ABB RobotStudio station: Pallet_Project.rspag

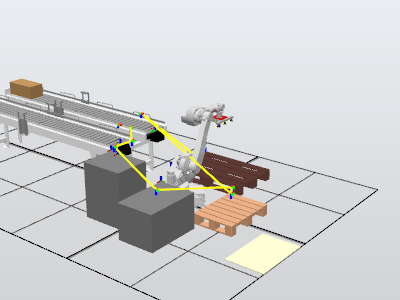
--- station ---
Station Pallet_Project (saved by RobotStudio 25.2.11220.0)
Controller Controler
  mechanical unit ROB_1: IRB1600_10_145__02, 6 joints, base frame (0, 0, 0) mm, rotated rx 0 ry 0 rz 135 deg
Layout (positions relative to the parent item):
  - IRB1600_10_145__02 [mechanism, from %ABB.RobotStudio.Models.IRB1600%\IRB1600_10_145_G_02.rslib] at (0, 0, 0) mm, rotated rx 0 ry 0 rz 135 deg; joint values [-2.2455, 0.5806, -0.4983, 0, 1.4885, 0.1107] (rad or m)
  - Half EPAL [part] at (-400, -600, 0) mm, rotated rx 0 ry 0 rz -90 deg, size 600 x 800 x 144 mm
  - ConveyorBox1 [part, from %ABB.RobotStudio.Models.Conveyors%\Conveyor Guide 400.rslib] at (150, 3660, 0) mm, rotated rx 0 ry 0 rz -90 deg
  - ConveyorBox2 [part, from %ABB.RobotStudio.Models.Conveyors%\Conveyor Guide 400.rslib] at (-550, 3660, 0) mm, rotated rx 0 ry 0 rz -90 deg
  - PalletizingVacuumTool [mechanism] at (1125, 125, 957.51) mm, rotated rx -180 ry 0 rz 180 deg
      TCP toolVacuum at (0, 0, 175) mm
      links: PalletizingVacuumTool
  - Box1 [part] at (338.5, 3410, 868) mm, size 249 x 499 x 200 mm
  - Box2 [part] at (-353.5, 3575, 868) mm, size 129 x 129 x 200 mm
  - EuroPallet [part, from Components\EuroPalletWood.rslib] at (1400, -600, 0) mm, rotated rx 0 ry 0 rz 90 deg
  - StackingTable [part], size 500 x 600 x 770 mm
  - LinerStand [part], size 800 x 540 x 500 mm
  - SC_Conveyor1 [smart component]
      signals: DO BoxArrived, DI EuroPalletReplaced, DO EuroPalletReplacedOut, DI EuroPalletFull
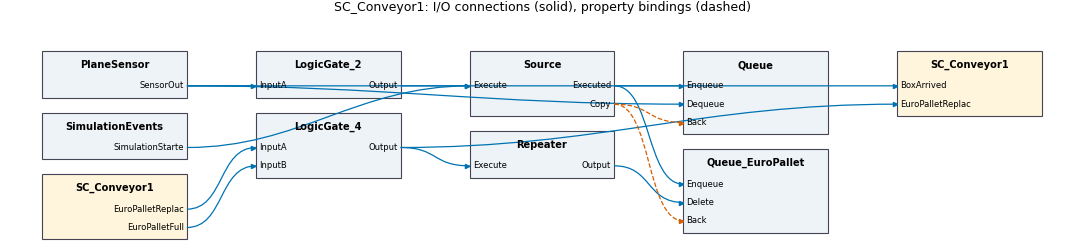
      connections:
        Source.Executed -> Queue.Enqueue
        PlaneSensor.SensorOut -> Queue.Dequeue
        PlaneSensor.SensorOut -> SC_Conveyor1.BoxArrived
        PlaneSensor.SensorOut -> LogicGate_2.InputA
        Source.Executed -> Queue_EuroPallet.Enqueue
        LogicGate_2.Output -> Source.Execute
        SimulationEvents.SimulationStarted -> Source.Execute
        SC_Conveyor1.EuroPalletReplaced -> LogicGate_4.InputA
        SC_Conveyor1.EuroPalletFull -> LogicGate_4.InputB
        LogicGate_4.Output -> Repeater.Execute
        LogicGate_4.Output -> SC_Conveyor1.EuroPalletReplacedOut
        Repeater.Output -> Queue_EuroPallet.Delete
        Source.Copy => Queue.Back
        Source.Copy => Queue_EuroPallet.Back
    - Source [smart component, from Components\Source.rslib]
        properties: Source=Box1; Copy=(none); Parent=(none); Position=[0.3385 3.39 0.868]; Orientation=[0 0 0]; Transient=true; PhysicsBehavior=-1
    - Queue [smart component, from Components\Queue.rslib]
        properties: Back=(none); Front=(none); Queue={81e52df3-1f77-4299-ba2a-6414327be985};{435d0d6d-d79b-44d3-acea-fe52ef949857};{8436b295-f8bf-4107-9481-0b8da08c6045};{6da8449d-009c-4835-8de1-a31c03bf24d8};{c517003d-8767-4c4a-bff9-7cbe8e804e1a};{f09c25fa-2584-409c-84e2-e14a50677c13};{130e9f86-ac44-4070-b92e-1e55d896aa7b};{906d2277-e14e-41d7-b5ad-7fe71654f1ef};{c971c019-2e6c-4537-9b43-f56770b68a66};{5740a0fa-eee5-4cb0-a52c-79e90074768b};{0e505042-845a-40e7-8904-6deb6f228de7};{2ef81a46-8090-4cc3-a468-447f4544bad1};{dd80a3b0-d0cd-4f2f-9600-d92ba7686845};{3b519026-604d-4377-8cfe-ae9118f60529}; NumberOfObjects=1
    - LinearMover [smart component, from Components\LinearMover.rslib]
        properties: Object=Queue; Direction=[0 -0.001 0]; Speed=0.25; Reference=Global; ReferenceObject=(none)
    - PlaneSensor [smart component, from Components\PlaneSensor.rslib]
        properties: Origin=[0.1885 0.675 0.788]; Axis1=[0.3 0 0]; Axis2=[0 0 0.01]; Tag=(none); SenseMultiple=false; SensedPart=(none)
      - _sensorPart_ [part], size 300 x 0 x 10 mm
    - LogicGate_2 [smart component, from Components\LogicGate.rslib]
        properties: Operator=NOT; Delay=0
    - SimulationEvents [smart component, from Components\SimulationEvents.rslib]
    - Queue_EuroPallet [smart component, from Components\Queue.rslib]
        properties: Back=(none); Front=(none); Queue={2ef81a46-8090-4cc3-a468-447f4544bad1};{dd80a3b0-d0cd-4f2f-9600-d92ba7686845};{3b519026-604d-4377-8cfe-ae9118f60529}; NumberOfObjects=3
    - LogicGate_4 [smart component, from Components\LogicGate.rslib]
        properties: Operator=AND; Delay=0
    - Repeater [smart component, from Components\Repeater.rslib]
        properties: Count=12
  - SC_Gripper [smart component]
      signals: DI Grip
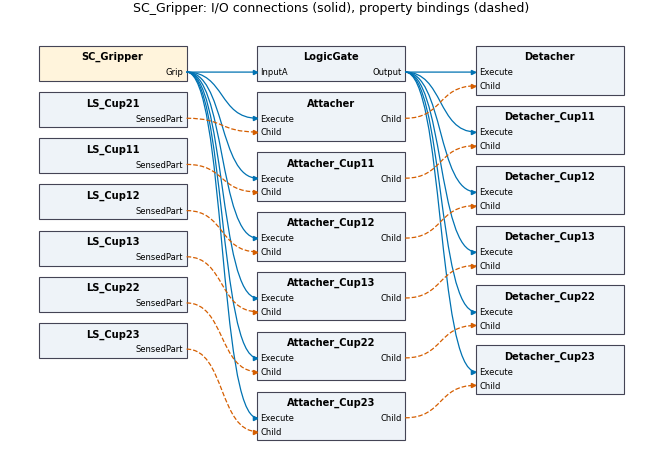
      connections:
        SC_Gripper.Grip -> Attacher.Execute
        SC_Gripper.Grip -> LogicGate.InputA
        LogicGate.Output -> Detacher.Execute
        SC_Gripper.Grip -> Attacher_Cup11.Execute
        LogicGate.Output -> Detacher_Cup11.Execute
        SC_Gripper.Grip -> Attacher_Cup12.Execute
        LogicGate.Output -> Detacher_Cup12.Execute
        SC_Gripper.Grip -> Attacher_Cup13.Execute
        LogicGate.Output -> Detacher_Cup13.Execute
        SC_Gripper.Grip -> Attacher_Cup22.Execute
        LogicGate.Output -> Detacher_Cup22.Execute
        SC_Gripper.Grip -> Attacher_Cup23.Execute
        LogicGate.Output -> Detacher_Cup23.Execute
        LS_Cup21.SensedPart => Attacher.Child
        Attacher.Child => Detacher.Child
        LS_Cup11.SensedPart => Attacher_Cup11.Child
        Attacher_Cup11.Child => Detacher_Cup11.Child
        LS_Cup12.SensedPart => Attacher_Cup12.Child
        Attacher_Cup12.Child => Detacher_Cup12.Child
        LS_Cup13.SensedPart => Attacher_Cup13.Child
        Attacher_Cup13.Child => Detacher_Cup13.Child
        LS_Cup22.SensedPart => Attacher_Cup22.Child
        Attacher_Cup22.Child => Detacher_Cup22.Child
        LS_Cup23.SensedPart => Attacher_Cup23.Child
        Attacher_Cup23.Child => Detacher_Cup23.Child
    - LS_Cup21 [smart component, from Components\LineSensor.rslib] at (375, 125, -163.99) mm, rotated rx 0 ry 0 rz -135 deg
        properties: Start=[-0.597509982704304 0.689429996191639 0.956499992313755]; End=[-0.597509981617333 0.689429995104668 0.924499992313755]; Length=0.032; Radius=0.00331491712707182; Tag=(none); SenseMultiple=false; SensedPart=(none); SensedPoint=[0 0 0]
      - _sensorPart_ [part], size 6.4 x 6.4 x 32 mm
    - Attacher [smart component, from Components\Attacher.rslib]
        properties: Parent=PalletizingVacuumTool; Flange=0; Child=(none); Mount=false; Offset=[0 0 0]; Orientation=[0 0 0]
    - Detacher [smart component, from Components\Detacher.rslib]
        properties: Child=(none); KeepPosition=true
    - LogicGate [smart component, from Components\LogicGate.rslib]
        properties: Operator=NOT; Delay=0
    - LS_Cup11 [smart component, from Components\LineSensor.rslib] at (375, 125, -163.99) mm, rotated rx 0 ry 0 rz -135 deg
        properties: Start=[-0.68943 0.59751 0.9565]; End=[-0.68943 0.59751 0.9245]; Length=0.032; Radius=0.00331; Tag=(none); SenseMultiple=false; SensedPart=(none); SensedPoint=[0 0 0]
      - _sensorPart_ [part], size 6.6 x 6.6 x 32 mm
    - LS_Cup12 [smart component, from Components\LineSensor.rslib] at (375, 125, -163.99) mm, rotated rx 0 ry 0 rz -135 deg
        properties: Start=[-0.57629 0.48437 0.9565]; End=[-0.57629 0.48437 0.9245]; Length=0.032; Radius=0.00331; Tag=(none); SenseMultiple=false; SensedPart=(none); SensedPoint=[0 0 0]
      - _sensorPart_ [part], size 6.6 x 6.6 x 32 mm
    - LS_Cup13 [smart component, from Components\LineSensor.rslib] at (375, 125, -163.99) mm, rotated rx 0 ry 0 rz -135 deg
        properties: Start=[-0.46315 0.37123 0.9565]; End=[-0.46315 0.37123 0.9245]; Length=0.032; Radius=0.00331; Tag=(none); SenseMultiple=false; SensedPart=(none); SensedPoint=[0 0 0]
      - _sensorPart_ [part], size 6.6 x 6.6 x 32 mm
    - LS_Cup22 [smart component, from Components\LineSensor.rslib] at (375, 125, -163.99) mm, rotated rx 0 ry 0 rz -135 deg
        properties: Start=[-0.48437 0.57629 0.9565]; End=[-0.48437 0.57629 0.9245]; Length=0.032; Radius=0.00331; Tag=(none); SenseMultiple=false; SensedPart=(none); SensedPoint=[0 0 0]
      - _sensorPart_ [part], size 6.6 x 6.6 x 32 mm
    - LS_Cup23 [smart component, from Components\LineSensor.rslib] at (375, 125, -163.99) mm, rotated rx 0 ry 0 rz -135 deg
        properties: Start=[-0.37123 0.46315 0.9565]; End=[-0.37123 0.46315 0.9245]; Length=0.032; Radius=0.00331; Tag=(none); SenseMultiple=false; SensedPart=(none); SensedPoint=[0 0 0]
      - _sensorPart_ [part], size 6.6 x 6.6 x 32 mm
    - Attacher_Cup11 [smart component, from Components\Attacher.rslib]
        properties: Parent=PalletizingVacuumTool; Flange=0; Child=(none); Mount=false; Offset=[0 0 0]; Orientation=[0 0 0]
    - Detacher_Cup11 [smart component, from Components\Detacher.rslib]
        properties: Child=(none); KeepPosition=true
    - Attacher_Cup12 [smart component, from Components\Attacher.rslib]
        properties: Parent=PalletizingVacuumTool; Flange=0; Child=(none); Mount=false; Offset=[0 0 0]; Orientation=[0 0 0]
    - Detacher_Cup12 [smart component, from Components\Detacher.rslib]
        properties: Child=(none); KeepPosition=true
    - Attacher_Cup13 [smart component, from Components\Attacher.rslib]
        properties: Parent=PalletizingVacuumTool; Flange=0; Child=(none); Mount=false; Offset=[0 0 0]; Orientation=[0 0 0]
    - Detacher_Cup13 [smart component, from Components\Detacher.rslib]
        properties: Child=(none); KeepPosition=true
    - Attacher_Cup22 [smart component, from Components\Attacher.rslib]
        properties: Parent=PalletizingVacuumTool; Flange=0; Child=(none); Mount=false; Offset=[0 0 0]; Orientation=[0 0 0]
    - Detacher_Cup22 [smart component, from Components\Detacher.rslib]
        properties: Child=(none); KeepPosition=true
    - Attacher_Cup23 [smart component, from Components\Attacher.rslib]
        properties: Parent=PalletizingVacuumTool; Flange=0; Child=(none); Mount=false; Offset=[0 0 0]; Orientation=[0 0 0]
    - Detacher_Cup23 [smart component, from Components\Detacher.rslib]
        properties: Child=(none); KeepPosition=true
  - SC_Conveyor2 [smart component]
      signals: DO BoxArrived, DI HalfPalletReplaced, DI HalfPalletFull, DO HalfPalletReplacedOut
      connections:
        Source.Executed -> Queue.Enqueue
        PlaneSensor.SensorOut -> Queue.Dequeue
        PlaneSensor.SensorOut -> SC_Conveyor2.BoxArrived
        PlaneSensor.SensorOut -> LogicGate.InputA
        SimulationEvents.SimulationStarted -> Source.Execute
        LogicGate.Output -> Source.Execute
        Repeater.Output -> Queue_HalfPallet.Delete
        SC_Conveyor2.HalfPalletReplaced -> LogicGate_5.InputA
        SC_Conveyor2.HalfPalletFull -> LogicGate_5.InputB
        LogicGate_5.Output -> Repeater.Execute
        LogicGate_5.Output -> SC_Conveyor2.HalfPalletReplacedOut
        Source.Executed -> Queue_HalfPallet.Enqueue
        Source.Copy => Queue.Back
        Source.Copy => Queue_HalfPallet.Back
    - Source [smart component, from Components\Source.rslib]
        properties: Source=Box2; Copy=(none); Parent=(none); Position=[-0.3535 3.575 0.868]; Orientation=[0 0 0]; Transient=true; PhysicsBehavior=-1
    - Queue [smart component, from Components\Queue.rslib]
        properties: Back=(none); Front=(none); Queue={9800cfb8-accd-4327-91e1-8f1786e05042};{c190d427-2878-4db8-b2be-214c692a7843};{b2a63077-10cd-4047-b774-a402e54bd5ce};{0cb034eb-9137-4204-8c4d-aa4d35edbbb2};{a2136454-01e3-48eb-803c-0c949220dd1f};{d1d29149-a959-4839-a5f8-05156c3e548d};{48c194bf-a44f-484f-bd23-34306ecfb550};{495763de-9b16-4c8d-83d3-4557bdb480a3};{abf2df07-53cd-488b-8dcb-fd67f1eb4dba}; NumberOfObjects=0
    - LinearMover [smart component, from Components\LinearMover.rslib]
        properties: Object=Queue; Direction=[0 -0.001 0]; Speed=0.25; Reference=Global; ReferenceObject=(none)
    - PlaneSensor [smart component, from Components\PlaneSensor.rslib]
        properties: Origin=[-0.5035 0.675 0.788]; Axis1=[0.3 0 0]; Axis2=[0 0 0.01]; Tag=(none); SenseMultiple=false; SensedPart=(none)
      - _sensorPart_ [part], size 300 x 0 x 10 mm
    - LogicGate [smart component, from Components\LogicGate.rslib]
        properties: Operator=NOT; Delay=0
    - SimulationEvents [smart component, from Components\SimulationEvents.rslib]
    - Queue_HalfPallet [smart component, from Components\Queue.rslib]
        properties: Back=(none); Front=(none); Queue={d5a67242-ef94-4595-a834-178362eb1d62};{353021ae-f387-47f5-aad2-fe3f1426ad48};{d78ca7a8-fd6f-498f-a8d6-0ea3578c76b0};{3356f02f-29aa-44c2-9ebf-5d29c5a600e5};{8f4d4553-4c1d-4056-aeb8-bca03c426780};{1a6d2d73-c05b-4390-90bb-4172aa34495b};{5c83e94b-c9dd-45e1-939f-1611cce13607};{08b3fadb-cba7-4510-a02f-3e66ae7e4329};{3ef4086a-d1f9-4a83-9755-3951cf9eaa00};{7bbd94bd-538e-428e-af81-32894a937116};{23a64fb5-90dc-4163-9a5d-a709f29cb737};{65ed0540-bcad-4628-84d7-59a3b9c76640};{b98fc11a-8ded-4a1c-bcf2-f2c76b1d1bd5};{5eac1296-3e35-4c81-a158-90d5fa5352fe};{05c4dc44-4e6c-4dc2-9677-a1940e3b3e4c};{d3d90d6c-55f3-41f9-ab59-03e6f986434c};{de9bd2e6-7614-4944-a633-7d4466c06302};{d5320c6f-757c-466b-aded-364807c4b01e};{23621476-4bd4-41d2-9f29-d7724955c74c};{817a93c2-45d8-40d3-ae92-600157ce3ee9};{243d6776-53f3-40e8-a26d-04ab6a776894};{7c17ee41-3d5e-4ce3-b2c1-8319b1484f6c};{7a467470-9a85-48d0-bfc9-40585f186b4a};{7fbfd87a-23fa-474d-b93a-b31788b7d83a};{49c53e7e-6fec-4cf6-ade2-eccfaa663d3f};{fd420bc1-af1d-47a6-a241-17656bc699f2};{1442cd0c-dbcc-4cc3-9371-290095dab2c2};{d4afd0ce-8611-4c71-934e-ce83a9ed8ab0};{4a599a5b-b82c-4c22-8dc8-b659788bcb6c};{af434e4d-6f74-4bd4-92e4-29d48b0c2391};{1d1a6925-ca0b-4280-b7e3-c3d429ecdeb1};{5f6f7c8a-25f7-4961-bc3d-06f26c3590e9};{0a446cc8-67bf-4709-be5a-1f56f3673959};{1af88ff7-cf78-4e6d-9326-b5fe289dfe55};{5a76c50a-250b-45d0-bcc3-a15c7678bea9};{ce2ad899-ab0c-4e8d-b6d7-b5ce0875e251};{41250e61-ba51-4579-939a-c1cb9538416c};{f048b52f-5fa1-4572-b32f-60b2a46e1837};{1087fd67-f502-4529-85a7-08891c247a62};{a8fcad14-50a7-40f1-a4f5-1777183cc2f1};{093bf0cb-478b-4d41-bc85-a01e6c4947d5};{ba12b4d4-5356-412c-9a5b-07d0d090cd25};{ef8538f7-904e-4b24-81ca-ce6b8f30748f};{1e7db033-e1a6-46cf-8960-0a3b92aa4569};{6ae3754e-0c7d-46a2-8cb0-0df03192a8af};{a9820d8c-191d-4cb3-b284-618a32150a08};{67edf359-12bc-49fc-a518-7b7d3cdaf041};{ad25e574-dc3f-4262-b019-213ebc35634b};{9ab4d7b7-70db-4a3c-b7ba-4ffa764225eb};{e3a4e5db-fe34-4e2c-bab2-f43d24e1bbe5};{2af16a20-02e3-4091-b49e-02ac578eafb8};{1fd54043-75f1-4856-9dc4-5fcdc28b2d30};{b3ff0692-c2c4-465f-bc5c-501c830a156d};{c5881555-d748-47b7-88bf-bb4395c5d677};{22d02747-187f-42da-b66b-aeac508d4faf};{4d19efbb-6ba8-4530-9818-c3b36a5b5e6d};{c26dfd74-1de5-480f-8d87-a956ac996da4};{800d2495-1f8a-4fba-a20e-307d73ad8d62};{4b542189-3f8e-408f-9294-fa7737ba2a1e};{b91039b3-272a-456d-b4ad-0c586638a480};{a02115cb-f377-4e0b-9fca-d98f58ac551d};{4b29cf1c-701e-48c2-bed8-74150284ae2a};{1a79b9b6-686e-4284-baae-745627c15955};{ca69f178-3ff4-4429-a57f-e75714190848};{2eeff9d0-5db0-4a2e-8983-6baf0d7612ee};{eb15173f-71b9-4843-b116-0fef5b8487ca};{f03858ea-60b5-4441-9128-abbe714a5bd1};{88a7fade-b898-403a-9912-eb07dfa3f617};{0c60aaed-4d54-4bbc-a941-b06aadfbebd1};{9800cfb8-accd-4327-91e1-8f1786e05042};{c190d427-2878-4db8-b2be-214c692a7843};{b2a63077-10cd-4047-b774-a402e54bd5ce};{0cb034eb-9137-4204-8c4d-aa4d35edbbb2};{a2136454-01e3-48eb-803c-0c949220dd1f};{d1d29149-a959-4839-a5f8-05156c3e548d};{48c194bf-a44f-484f-bd23-34306ecfb550};{495763de-9b16-4c8d-83d3-4557bdb480a3};{abf2df07-53cd-488b-8dcb-fd67f1eb4dba}; NumberOfObjects=32
    - Repeater [smart component, from Components\Repeater.rslib]
        properties: Count=72
    - LogicGate_5 [smart component, from Components\LogicGate.rslib]
        properties: Operator=AND; Delay=0
  - Liner_01 [part] at (-900, -2000, 0) mm, size 800 x 540 x 10 mm
  - SC_Liners [smart component]
      signals: DI LinersRefilled, DI LinerStackEmpty, DI PalletReplaced, DO LinersRefilledOut
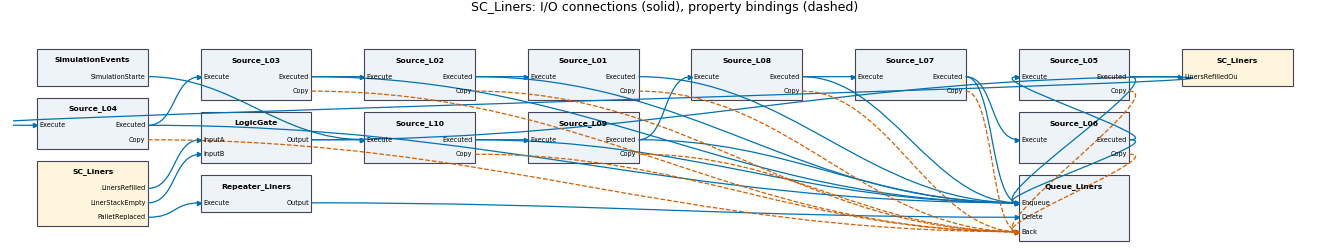
      connections:
        SimulationEvents.SimulationStarted -> Source_L10.Execute
        Source_L10.Executed -> Queue_Liners.Enqueue
        Source_L10.Executed -> Source_L09.Execute
        Source_L09.Executed -> Queue_Liners.Enqueue
        Source_L09.Executed -> Source_L08.Execute
        Source_L08.Executed -> Queue_Liners.Enqueue
        Source_L08.Executed -> Source_L07.Execute
        Source_L07.Executed -> Queue_Liners.Enqueue
        Source_L07.Executed -> Source_L06.Execute
        Source_L06.Executed -> Queue_Liners.Enqueue
        Source_L06.Executed -> Source_L05.Execute
        Source_L05.Executed -> Queue_Liners.Enqueue
        Source_L05.Executed -> Source_L04.Execute
        Source_L04.Executed -> Queue_Liners.Enqueue
        Source_L04.Executed -> Source_L03.Execute
        Source_L03.Executed -> Queue_Liners.Enqueue
        Source_L03.Executed -> Source_L02.Execute
        Source_L02.Executed -> Queue_Liners.Enqueue
        Source_L02.Executed -> Source_L01.Execute
        Source_L01.Executed -> Queue_Liners.Enqueue
        SC_Liners.LinersRefilled -> LogicGate.InputA
        SC_Liners.LinerStackEmpty -> LogicGate.InputB
        LogicGate.Output -> SC_Liners.LinersRefilledOut
        LogicGate.Output -> Source_L10.Execute
        SC_Liners.PalletReplaced -> Repeater_Liners.Execute
        Repeater_Liners.Output -> Queue_Liners.Delete
        Source_L10.Copy => Queue_Liners.Back
        Source_L09.Copy => Queue_Liners.Back
        Source_L08.Copy => Queue_Liners.Back
        Source_L07.Copy => Queue_Liners.Back
        Source_L06.Copy => Queue_Liners.Back
        Source_L05.Copy => Queue_Liners.Back
        Source_L04.Copy => Queue_Liners.Back
        Source_L03.Copy => Queue_Liners.Back
        Source_L02.Copy => Queue_Liners.Back
        Source_L01.Copy => Queue_Liners.Back
    - Source_L10 [smart component, from Components\Source.rslib]
        properties: Source=Liner_01; Copy=(none); Parent=(none); Position=[-1.3 -0.7 0.59]; Orientation=[0 0 0]; Transient=true; PhysicsBehavior=-1
    - Source_L09 [smart component, from Components\Source.rslib]
        properties: Source=Liner_01; Copy=(none); Parent=(none); Position=[-1.3 -0.7 0.58]; Orientation=[0 0 0]; Transient=true; PhysicsBehavior=-1
    - Queue_Liners [smart component, from Components\Queue.rslib]
        properties: Back=(none); Front=(none); Queue={20d974b6-189e-48d5-91a3-27801e75a2e3};{290c2d17-6faa-4c17-875c-80c899971b7e};{09f81150-e011-45c7-9a87-29c6d5ac92f7};{b296464f-7b57-4359-8933-3b585c425c6c};{a4bcdc79-e721-4592-ba3d-6f160afd2660};{d0cb2024-c7d0-4f62-9559-4447ca439c63};{f1537fa3-356e-4cfb-b79c-b3a3ef2d5a1a};{ade4e0be-57dc-4cbd-9040-6b29c36965ae};{068dc0fe-76cb-4174-b384-f9a97e7185e6};{74ebf040-bda5-45b9-9c71-05d8b50facaf};{455b281d-0163-4b9a-96ec-b3dbceeb94ec};{5721ff76-6329-4602-9dd2-421615ef1c3b}; NumberOfObjects=10
    - SimulationEvents [smart component, from Components\SimulationEvents.rslib]
    - Source_L08 [smart component, from Components\Source.rslib]
        properties: Source=Liner_01; Copy=(none); Parent=(none); Position=[-1.3 -0.7 0.57]; Orientation=[0 0 0]; Transient=true; PhysicsBehavior=-1
    - Source_L07 [smart component, from Components\Source.rslib]
        properties: Source=Liner_01; Copy=(none); Parent=(none); Position=[-1.3 -0.7 0.56]; Orientation=[0 0 0]; Transient=true; PhysicsBehavior=-1
    - Source_L06 [smart component, from Components\Source.rslib]
        properties: Source=Liner_01; Copy=(none); Parent=(none); Position=[-1.3 -0.7 0.55]; Orientation=[0 0 0]; Transient=true; PhysicsBehavior=-1
    - Source_L05 [smart component, from Components\Source.rslib]
        properties: Source=Liner_01; Copy=(none); Parent=(none); Position=[-1.3 -0.7 0.54]; Orientation=[0 0 0]; Transient=true; PhysicsBehavior=-1
    - Source_L04 [smart component, from Components\Source.rslib]
        properties: Source=Liner_01; Copy=(none); Parent=(none); Position=[-1.3 -0.7 0.53]; Orientation=[0 0 0]; Transient=true; PhysicsBehavior=-1
    - Source_L03 [smart component, from Components\Source.rslib]
        properties: Source=Liner_01; Copy=(none); Parent=(none); Position=[-1.3 -0.7 0.52]; Orientation=[0 0 0]; Transient=true; PhysicsBehavior=-1
    - Source_L02 [smart component, from Components\Source.rslib]
        properties: Source=Liner_01; Copy=(none); Parent=(none); Position=[-1.3 -0.7 0.51]; Orientation=[0 0 0]; Transient=true; PhysicsBehavior=-1
    - Source_L01 [smart component, from Components\Source.rslib]
        properties: Source=Liner_01; Copy=(none); Parent=(none); Position=[-1.3 -0.7 0.5]; Orientation=[0 0 0]; Transient=true; PhysicsBehavior=-1
    - LogicGate [smart component, from Components\LogicGate.rslib]
        properties: Operator=AND; Delay=0
    - Repeater_Liners [smart component, from Components\Repeater.rslib]
        properties: Count=2
Attachment: PalletizingVacuumTool is attached to IRB1600_10_145__02 / Link6
Attachment: LS_Cup21 is attached to PalletizingVacuumTool / PalletizingVacuumTool
Attachment: LS_Cup12 is attached to PalletizingVacuumTool / PalletizingVacuumTool
Attachment: LS_Cup13 is attached to PalletizingVacuumTool / PalletizingVacuumTool
Attachment: LS_Cup22 is attached to PalletizingVacuumTool / PalletizingVacuumTool
Attachment: LS_Cup23 is attached to PalletizingVacuumTool / PalletizingVacuumTool
Attachment: LS_Cup11 is attached to PalletizingVacuumTool / PalletizingVacuumTool
Collision set Conjunto de colisión_1: IRB1600_10_145__02, PalletizingVacuumTool against ConveyorBox1, ConveyorBox2, EuroPallet, Half EPAL, LinerStand, StackingTable, near miss 0.05 m
Station logic (signal -> signal, property => property):
  SC_Conveyor1.BoxArrived -> Controler.DI_Box1Arrived
  Controler.DO_Cup21 -> SC_Gripper.Grip
  SC_Conveyor2.BoxArrived -> Controler.DI_Box2Arrived
  SC_Conveyor1.EuroPalletReplacedOut -> Controler.DI_EuroPalletReplaced
  Controler.DO_EuroPalletFull -> SC_Conveyor1.EuroPalletFull
  Controler.DO_HalfPalletFull -> SC_Conveyor2.HalfPalletFull
  SC_Conveyor2.HalfPalletReplacedOut -> Controler.DI_HalfPalletReplaced
  Controler.DO_LinerStackEmpty -> SC_Liners.LinerStackEmpty
  SC_Liners.LinersRefilledOut -> Controler.DI_LinersRefilled
  SC_Conveyor2.HalfPalletReplacedOut -> SC_Liners.PalletReplaced
Targets, tools, work objects and paths stored in the station and not in the controller backup, written as RAPID:
! task T_ROB1
MODULE PalletProgram
  PROC Path_10()
    MoveL PickConveyor2,v1000,z100,toolVacuum\WObj:=wobjConveyor2;
    MoveL PlaceTable,v1000,z100,toolVacuum\WObj:=wobjTable;
    MoveL PickTableStack,v1000,z100,toolVacuum\WObj:=wobjTable;
    MoveL PickLiner,v1000,z100,toolVacuum\WObj:=wobjLinerStack;
    MoveL PlaceHalfPallet,v1000,z100,toolVacuum\WObj:=wobjHalfPallet;
    MoveL PlaceLiner,v1000,z100,toolVacuum\WObj:=wobjHalfPallet;
    MoveL PickConveyor1,v1000,z100,toolVacuum\WObj:=wobjConveyor1;
    MoveL PlaceEuroRow2,v1000,z100,toolVacuum\WObj:=wobjEuroPallet;
    MoveL PlaceEuroRow4,v1000,z100,toolVacuum\WObj:=wobjEuroPallet;
  ENDPROC
ENDMODULE


--- Controller Data/Controler/RAPID/TASK1/PROGMOD/CalibData.mod ---
MODULE CalibData
    !-----------------------------------------------------------------------
	! Tools and work object
	!-----------------------------------------------------------------------
    TASK PERS wobjdata wobjEuroPallet:=[FALSE,TRUE,"",[[600,600,144],[0.707106781,0,0,-0.707106781]],[[0,0,0],[1,0,0,0]]];
    TASK PERS wobjdata wobjHalfPallet:=[FALSE,TRUE,"",[[400,-600,144],[0,0,0,1]],[[0,0,0],[1,0,0,0]]];
    TASK PERS wobjdata wobjConveyor1:=[FALSE,TRUE,"",[[338.5,670,768],[0.707106781,0,0,0.707106781]],[[0,0,0],[1,0,0,0]]];
    TASK PERS wobjdata wobjConveyor2:=[FALSE,TRUE,"",[[-353.5,670,768],[0.707106781,0,0,0.707106781]],[[0,0,0],[1,0,0,0]]];
    TASK PERS wobjdata wobjTable:=[FALSE,TRUE,"",[[-600,600,770],[0,0,0,1]],[[55,170,0],[1,0,0,0]]];
    TASK PERS wobjdata wobjLinerStack:=[FALSE,TRUE,"",[[-500,-160,500],[0,0,0,1]],[[0,0,0],[1,0,0,0]]];
    TASK PERS tooldata toolVacuum:=[TRUE,[[0,0,175],[1,0,0,0]],[1,[0,0,1],[1,0,0,0],0,0,0]];
    ! toolVacuum: mass and CoG are provisional (1 kg), to be estimated

    !-----------------------------------------------------------------------
	! Load data
	!-----------------------------------------------------------------------
    ! Payloads: CoG relative to the TCP of toolVacuum; inertia set to 0 (point mass) until confirmed
    TASK PERS loaddata loadBox1:=[2,[0,0,100],[1,0,0,0],0,0,0];
    ! Box 2 is picked with one corner cup (x=-160, y=-100); on the table fill rows ascending Y, each row descending X
    TASK PERS loaddata loadBox2:=[0.4,[-160,-100,100],[1,0,0,0],0,0,0];
    ! 3x2 stack of box 2 (390 x 260 x 200 mm, 6 x 0.4 kg)
    TASK PERS loaddata loadBox2Stack:=[2.4,[0,0,100],[1,0,0,0],0,0,0];
    ! Liner: corrugated cardboard, 0.8 x 0.54 x 0.01 m3 x 120 kg/m3 = 0.52 kg
    TASK PERS loaddata loadLiner:=[0.52,[0,0,5],[1,0,0,0],0,0,0];
ENDMODULE

--- Controller Data/Controler/RAPID/TASK1/PROGMOD/PalletProgram.mod ---
MODULE PalletProgram

    !***********************************************************************
    ! Industrial Robotics and Offline Programming G1F - University of Skovde
    ! Offline programming project: Pallet Project - Group 2 (JMPM)
    ! Authors: Peru Mendivil and Joaquin Moreno
    ! Robot :   ABB IRB 1600-10/1.45, IRC5 RobotWare 6.13.02 (RobotStudio 2025)
    ! Tool  :   toolVacuum, vacuum gripper with 6 cups (one valve per cup)
    ! Date:    2026-10-30
    !
    ! The robot palletizes two products coming on two conveyors.
    ! Box 1 goes from conveyor 1 to the Euro pallet: 4-2 pattern,
    ! 2 layers (12 boxes). Box 2 goes from conveyor 2 to the stacking
    ! table, where a 3x2 block is formed. The block is then moved to the
    ! half pallet: 2x2 blocks per layer, 3 layers (72 boxes), with a liner
    ! after layers 1 and 2. When both conveyors have a box, the robot
    ! alternates box 1 and box 2. A full pallet is replaced by the operator
    ! from outside the fence, and the robot keeps working with the other
    ! product. With the half pallet full, one block can still be finished
    ! on the table, and it waits there. If the liner stack is empty, the
    ! robot keeps working until a liner is needed; then box 2 waits until
    ! the operator refills the stack.
    !
    ! Structure: Main is a state machine (grafcet). It initialises the
    ! signals and then decides each cycle which box to handle, from the
    ! conveyor sensors, the full-pallet flags and the last box handled.
    ! Each product has its own routine with a finite-state machine for
    ! the place positions. Every place position is calculated with Offs
    ! from one base target per station. ApproachPoint does every
    ! pick/place: approach, vacuum on/off and GripLoad. Work objects,
    ! tool and loads are in the module CalibData.
    ! The operator buttons (pallet replaced, liners refilled) are read
    ! with interrupts (TRAP), so a short press is never lost.
    !
    ! Naming: VAR, PERS and parameters in camelCase (can change);
    ! CONST, PROC, FUNC and MODULE in PascalCase (fixed).
    !***********************************************************************

    !-----------------------------------------------------------------------
    ! Base targets
    !-----------------------------------------------------------------------
    CONST jointtarget Home:=[[0,0,0,0,90,0],[9E+09,9E+09,9E+09,9E+09,9E+09,9E+09]];

    ! Box 1
    CONST robtarget PickConveyor1:=[[249.5,0,200],[0,0,1,0],[0,0,0,0],[9E+09,9E+09,9E+09,9E+09,9E+09,9E+09]];
    CONST robtarget PlaceEuroRow4:=[[225,525,200],[0,-0.707106781,0.707106781,0],[-2,0,0,0],[9E+09,9E+09,9E+09,9E+09,9E+09,9E+09]];
    CONST robtarget PlaceEuroRow2:=[[350,150,200],[0,1,0,0],[-2,0,-1,0],[9E+09,9E+09,9E+09,9E+09,9E+09,9E+09]];

    ! Box 2
    CONST robtarget PickConveyor2:=[[-35.5,-160,200],[0,-0.707106781,0.707106781,0],[0,0,0,0],[9E+09,9E+09,9E+09,9E+09,9E+09,9E+09]];
    CONST robtarget PlaceTable:=[[-95,165,200],[0,0,1,0],[0,0,0,0],[9E+09,9E+09,9E+09,9E+09,9E+09,9E+09]];
    CONST robtarget PickTableStack:=[[195,130,200],[0,0,1,0],[0,0,0,0],[9E+09,9E+09,9E+09,9E+09,9E+09,9E+09]];
    CONST robtarget PlaceHalfPallet:=[[205,170,200],[0,0,1,0],[0,0,0,0],[9E+09,9E+09,9E+09,9E+09,9E+09,9E+09]];

    ! Liners
    CONST robtarget PickLiner:=[[400,270,100],[0,0,1,0],[0,0,0,0],[9E+09,9E+09,9E+09,9E+09,9E+09,9E+09]];
    CONST robtarget PlaceLiner:=[[400,300,210],[0,0,1,0],[0,0,0,0],[9E+09,9E+09,9E+09,9E+09,9E+09,9E+09]];

    !-----------------------------------------------------------------------
    ! Speeds and heights
    !-----------------------------------------------------------------------
    CONST speeddata TransitSpeed:=v1000;
    CONST speeddata ApproachSpeed:=v300;

    ! Height of every station (world)
    CONST num ConveyorsHeight:=768;
    CONST num TableHeight:=770;
    CONST num LinerStandHeight:=500;
    CONST num EuroPalletHeight:=144;
    CONST num HalfPalletHeight:=144;

    CONST num Box1Height:=200;
    CONST num Box2Height:=200;

    ! Heights for the approach points
    CONST num TransitHeight:=1100;
    CONST num PalletOffsetHeight:=250;
    CONST num MinApproachHeight:=250;

    ! Station identifiers for ApproachHeight
    CONST num StationConveyor1:=1;
    CONST num StationConveyor2:=2;
    CONST num StationTable:=3;
    CONST num StationLinerStand:=4;
    CONST num StationHalfPallet:=5;
    CONST num StationEuroPallet:=6;

    !-----------------------------------------------------------------------
    ! Vacuum gripper
    !-----------------------------------------------------------------------
    CONST num VacuumTime:=1;
    CONST bool CupsAllOn{6}:=[TRUE,TRUE,TRUE,TRUE,TRUE,TRUE];
    CONST bool CupsAllOff{6}:=[FALSE,FALSE,FALSE,FALSE,FALSE,FALSE];
    CONST bool CupsBox2On{6}:=[FALSE,FALSE,FALSE,TRUE,FALSE,FALSE];
    VAR bool cupsState{6}:=[FALSE,FALSE,FALSE,FALSE,FALSE,FALSE];
    VAR signaldo cupSignals{6};

    !-----------------------------------------------------------------------
    ! Box selection
    !-----------------------------------------------------------------------
    CONST num Box1:=1;
    CONST num Box2:=2;
    ! Last box handled, to alternate box 1 and box 2
    VAR num lastBox:=Box2;

    !-----------------------------------------------------------------------
    ! Box 1 state machine parameters and variables
    !-----------------------------------------------------------------------
    CONST num Box1Pos1:=1;
    CONST num Box1Pos2:=2;
    CONST num Box1Pos3:=3;
    CONST num Box1Pos4:=4;
    CONST num Box1Pos5:=5;
    CONST num Box1LastPos:=6;
    CONST num Box1MaxLayers:=2;
    ! Distance between boxes in the row of 4 and in the row of 2
    CONST num EuroRow4Offset:=250;
    CONST num EuroRow2Offset:=500;

    VAR num box1State:=1;
    VAR num box1Layer:=1;
    VAR bool euroPalletFull:=FALSE;

    ! Euro pallet replaced by the operator: interrupt and flag set by the TRAP
    VAR intnum euroReplacedInt;
    VAR bool euroPalletReplaced:=FALSE;

    !-----------------------------------------------------------------------
    ! Box 2 state machine parameters and variables (table)
    !-----------------------------------------------------------------------
    CONST num Box2Pos1:=1;
    CONST num Box2Pos2:=2;
    CONST num Box2Pos3:=3;
    CONST num Box2Pos4:=4;
    CONST num Box2Pos5:=5;
    CONST num Box2LastPos:=6;
    ! Distance between boxes 2 on the table
    CONST num Box2Offset:=130;

    VAR num box2State:=1;
    VAR bool tableFull:=FALSE;

    !-----------------------------------------------------------------------
    ! TransferStack parameters and variables (half pallet)
    !-----------------------------------------------------------------------
    CONST num BlockPos1:=1;
    CONST num BlockPos2:=2;
    CONST num BlockPos3:=3;
    CONST num BlockPos4:=4;
    CONST num Box2MaxLayers:=3;
    ! Distance between 3x2 blocks on the half pallet
    CONST num BlockOffsetX:=3*Box2Offset;
    CONST num BlockOffsetY:=2*Box2Offset;

    VAR num blockState:=1;
    VAR num box2Layer:=1;
    VAR bool halfPalletFull:=FALSE;

    ! Half pallet replaced by the operator: interrupt and flag set by the TRAP
    VAR intnum halfReplacedInt;
    VAR bool halfPalletReplaced:=FALSE;

    !-----------------------------------------------------------------------
    ! Liners parameters and variables
    !-----------------------------------------------------------------------
    CONST num TotalLiners:=10;
    CONST num LinerHeight:=10;

    VAR num linersLeft:=TotalLiners;
    ! Liner stack empty: warning to the operator, the robot keeps working
    VAR bool linerStackEmpty:=FALSE;
    ! Layer complete but the liner stack is empty: box 2 waits for the refill
    VAR bool linerMissing:=FALSE;

    ! Liners refilled by the operator: interrupt and flag set by the TRAP
    VAR intnum linersRefilledInt;
    VAR bool linersRefilled:=FALSE;

    !-----------------------------------------------------------------------
    ! Main: choose the box and check the operator signals
    !-----------------------------------------------------------------------
    PROC Main()

        InitSignals;
        VacuumControl CupsAllOff;
        SetDO DO_EuroPalletFull,0;
        SetDO DO_HalfPalletFull,0;
        SetDO DO_LinerStackEmpty,0;
        ! Connect an interrupt to DI_EuroPalletReplaced: EuroPalletReplacedTrap runs on every rising edge
        IDelete euroReplacedInt;
        CONNECT euroReplacedInt WITH EuroPalletReplacedTrap;
        ISignalDI DI_EuroPalletReplaced,1,euroReplacedInt;
        ! Connect an interrupt to DI_HalfPalletReplaced: HalfPalletReplacedTrap runs on every rising edge
        IDelete halfReplacedInt;
        CONNECT halfReplacedInt WITH HalfPalletReplacedTrap;
        ISignalDI DI_HalfPalletReplaced,1,halfReplacedInt;
        ! Connect an interrupt to DI_LinersRefilled: LinersRefilledTrap runs on every rising edge
        IDelete linersRefilledInt;
        CONNECT linersRefilledInt WITH LinersRefilledTrap;
        ISignalDI DI_LinersRefilled,1,linersRefilledInt;
        GripLoad load0;
        MoveAbsJ Home,v100,fine,toolVacuum;

        WHILE TRUE DO

            ! Alternate box 1 and box 2 when both are ready
            IF Box1Ready() AND ((NOT Box2Ready()) OR lastBox=Box2) THEN
                ProcessBox1;
            ELSEIF Box2Ready() THEN
                ProcessBox2;
            ENDIF

            ! Euro pallet replaced (flag set by the TRAP): back to layer 1
            IF euroPalletReplaced THEN
                euroPalletReplaced:=FALSE;
                box1Layer:=1;
                ! Not necessary but safe
                box1State:=Box1Pos1;
                euroPalletFull:=FALSE;
            ENDIF

            ! Half pallet replaced (flag set by the TRAP): layer 1 first, then the waiting block
            IF halfPalletReplaced THEN
                halfPalletReplaced:=FALSE;
                box2Layer:=1;
                blockState:=BlockPos1;
                halfPalletFull:=FALSE;
                IF tableFull THEN
                    TransferStack;
                    tableFull:=FALSE;
                ENDIF
            ENDIF

            ! Liners refilled (flag set by the TRAP): reload the counter, then the missing liner and the waiting block
            IF linersRefilled THEN
                linersRefilled:=FALSE;
                linersLeft:=TotalLiners;
                linerStackEmpty:=FALSE;
                IF linerMissing THEN
                    linerMissing:=FALSE;
                    PlaceLayerLiner;
                    IF tableFull THEN
                        TransferStack;
                        tableFull:=FALSE;
                    ENDIF
                ENDIF
            ENDIF
            WaitTime 0.1;
        ENDWHILE
    ENDPROC

    !-----------------------------------------------------------------------
    ! Interrupts: operator buttons (pallet replaced, liners refilled)
    !-----------------------------------------------------------------------
    TRAP EuroPalletReplacedTrap
        ! Only considered if the pallet is already full to prevent false positives
        IF euroPalletFull THEN
            ! Light off at once, even while the robot moves: the operator instantly sees the press was accepted
            SetDO DO_EuroPalletFull,0;
            ! Main sets layer 1 when the robot is free (no motion in a TRAP)
            euroPalletReplaced:=TRUE;
        ENDIF
    ENDTRAP

    TRAP HalfPalletReplacedTrap
        ! Only considered if the pallet is already full to prevent false positives
        IF halfPalletFull THEN
            ! Light off at once, even while the robot moves: the operator instantly sees the press was accepted
            SetDO DO_HalfPalletFull,0;
            ! Main sets layer 1 and moves the waiting block (no motion in a TRAP)
            halfPalletReplaced:=TRUE;
        ENDIF
    ENDTRAP

    TRAP LinersRefilledTrap
        ! Only if the stack is empty, to prevent false positives
        IF linerStackEmpty THEN
            ! Light off at once, even while the robot moves: the operator instantly sees the press was accepted
            SetDO DO_LinerStackEmpty,0;
            ! Main reloads the counter, then places the missing liner and block (no motion in a TRAP)
            linersRefilled:=TRUE;
        ENDIF
    ENDTRAP

    !-----------------------------------------------------------------------
    ! Box ready to be handled
    !-----------------------------------------------------------------------
    FUNC bool Box1Ready()
        ! Box 1 waiting on conveyor 1 and room on the Euro pallet
        RETURN (DI_Box1Arrived=1) AND (NOT euroPalletFull);
    ENDFUNC

    FUNC bool Box2Ready()
        ! Box 2 waiting on conveyor 2 and room on the table
        RETURN (DI_Box2Arrived=1) AND (NOT tableFull);
    ENDFUNC

    !-----------------------------------------------------------------------
    ! Box 1 state machine: conveyor 1 to the Euro pallet
    !-----------------------------------------------------------------------
    PROC ProcessBox1()
        ! Z of the current layer on the Euro pallet
        VAR num layerZ;

        ApproachPoint PickConveyor1,wobjConveyor1,CupsAllOn,loadBox1,ApproachHeight(StationConveyor1);

        layerZ:=(box1Layer-1)*Box1Height;
        TEST box1State
        CASE Box1Pos1:
            ApproachPoint Offs(PlaceEuroRow4,0,0,layerZ),wobjEuroPallet,CupsAllOff,load0,ApproachHeight(StationEuroPallet);
            box1State:=Box1Pos2;
        CASE Box1Pos2:
            ApproachPoint Offs(PlaceEuroRow4,EuroRow4Offset,0,layerZ),wobjEuroPallet,CupsAllOff,load0,ApproachHeight(StationEuroPallet);
            box1State:=Box1Pos3;
        CASE Box1Pos3:
            ApproachPoint Offs(PlaceEuroRow4,2*EuroRow4Offset,0,layerZ),wobjEuroPallet,CupsAllOff,load0,ApproachHeight(StationEuroPallet);
            box1State:=Box1Pos4;
        CASE Box1Pos4:
            ApproachPoint Offs(PlaceEuroRow4,3*EuroRow4Offset,0,layerZ),wobjEuroPallet,CupsAllOff,load0,ApproachHeight(StationEuroPallet);
            box1State:=Box1Pos5;
        CASE Box1Pos5:
            ApproachPoint Offs(PlaceEuroRow2,0,0,layerZ),wobjEuroPallet,CupsAllOff,load0,ApproachHeight(StationEuroPallet);
            box1State:=Box1LastPos;
        CASE Box1LastPos:
            ApproachPoint Offs(PlaceEuroRow2,EuroRow2Offset,0,layerZ),wobjEuroPallet,CupsAllOff,load0,ApproachHeight(StationEuroPallet);
            IF box1Layer=Box1MaxLayers THEN
                euroPalletFull:=TRUE;
                SetDO DO_EuroPalletFull,1;
            ELSE
                Incr box1Layer;
            ENDIF
            box1State:=Box1Pos1;
        DEFAULT:
            box1State:=Box1Pos1;
        ENDTEST
        lastBox:=Box1;
    ENDPROC

    !-----------------------------------------------------------------------
    ! Box 2 state machine: conveyor 2 to the table
    !-----------------------------------------------------------------------
    PROC ProcessBox2()

        ApproachPoint PickConveyor2,wobjConveyor2,CupsBox2On,loadBox2,ApproachHeight(StationConveyor2);

        ! Far row (y=130) first and x from high to low: the box carried never crosses the boxes already placed
        TEST box2State
        CASE Box2Pos1:
            ApproachPoint Offs(PlaceTable,2*Box2Offset,Box2Offset,0),wobjTable,CupsAllOff,load0,ApproachHeight(StationTable);
            box2State:=Box2Pos2;
        CASE Box2Pos2:
            ApproachPoint Offs(PlaceTable,Box2Offset,Box2Offset,0),wobjTable,CupsAllOff,load0,ApproachHeight(StationTable);
            box2State:=Box2Pos3;
        CASE Box2Pos3:
            ApproachPoint Offs(PlaceTable,0,Box2Offset,0),wobjTable,CupsAllOff,load0,ApproachHeight(StationTable);
            box2State:=Box2Pos4;
        CASE Box2Pos4:
            ApproachPoint Offs(PlaceTable,2*Box2Offset,0,0),wobjTable,CupsAllOff,load0,ApproachHeight(StationTable);
            box2State:=Box2Pos5;
        CASE Box2Pos5:
            ApproachPoint Offs(PlaceTable,Box2Offset,0,0),wobjTable,CupsAllOff,load0,ApproachHeight(StationTable);
            box2State:=Box2LastPos;
        CASE Box2LastPos:
            ApproachPoint Offs(PlaceTable,0,0,0),wobjTable,CupsAllOff,load0,ApproachHeight(StationTable);
            IF halfPalletFull OR linerMissing THEN
                tableFull:=TRUE;
            ELSE
                TransferStack;
            ENDIF
            box2State:=Box2Pos1;
        DEFAULT:
            box2State:=Box2Pos1;
        ENDTEST
        lastBox:=Box2;
    ENDPROC

    !-----------------------------------------------------------------------
    ! Box 2: move the 3x2 block from the table to the half pallet
    !-----------------------------------------------------------------------
    PROC TransferStack()
        ! Z of the current layer on the half pallet (block and liner)
        VAR num layerZ;

        ! Pick all 6 boxes 2
        ApproachPoint PickTableStack,wobjTable,CupsAllOn,loadBox2Stack,ApproachHeight(StationTable);

        ! Place group of boxes
        layerZ:=HalfPalletLayerZ();
        TEST blockState
        CASE BlockPos1:
            ApproachPoint Offs(PlaceHalfPallet,0,BlockOffsetY,layerZ),wobjHalfPallet,CupsAllOff,load0,ApproachHeight(StationHalfPallet);
            blockState:=BlockPos2;
        CASE BlockPos2:
            ApproachPoint Offs(PlaceHalfPallet,BlockOffsetX,BlockOffsetY,layerZ),wobjHalfPallet,CupsAllOff,load0,ApproachHeight(StationHalfPallet);
            blockState:=BlockPos3;
        CASE BlockPos3:
            ApproachPoint Offs(PlaceHalfPallet,0,0,layerZ),wobjHalfPallet,CupsAllOff,load0,ApproachHeight(StationHalfPallet);
            blockState:=BlockPos4;
        CASE BlockPos4:
            ApproachPoint Offs(PlaceHalfPallet,BlockOffsetX,0,layerZ),wobjHalfPallet,CupsAllOff,load0,ApproachHeight(StationHalfPallet);
            IF box2Layer=Box2MaxLayers THEN
                halfPalletFull:=TRUE;
                SetDO DO_HalfPalletFull,1;
            ELSEIF linerStackEmpty THEN
                linerMissing:=TRUE;
            ELSE
                PlaceLayerLiner;
            ENDIF
            blockState:=BlockPos1;
        DEFAULT:
            blockState:=BlockPos1;
        ENDTEST
    ENDPROC

    !-----------------------------------------------------------------------
    ! Liner on the layer just finished, then the next layer starts
    !-----------------------------------------------------------------------
    PROC PlaceLayerLiner()
        ApproachPoint Offs(PickLiner,0,0,-(TotalLiners-linersLeft)*LinerHeight),wobjLinerStack,CupsAllOn,loadLiner,ApproachHeight(StationLinerStand);
        ApproachPoint Offs(PlaceLiner,0,0,HalfPalletLayerZ()),wobjHalfPallet,CupsAllOff,load0,ApproachHeight(StationHalfPallet);
        Incr box2Layer;
        Decr linersLeft;
        IF linersLeft=0 THEN
            linerStackEmpty:=TRUE;
            SetDO DO_LinerStackEmpty,1;
        ENDIF
    ENDPROC

    !-----------------------------------------------------------------------
    ! Z of the current layer on the half pallet (block and liner)
    !-----------------------------------------------------------------------
    FUNC num HalfPalletLayerZ()
        ! One liner under every layer except the first one
        RETURN (box2Layer-1)*(Box2Height+LinerHeight);
    ENDFUNC

    !-----------------------------------------------------------------------
    ! Pick or place at a target: approach, vacuum, GripLoad and go up
    !-----------------------------------------------------------------------
    PROC ApproachPoint(robtarget target,PERS wobjdata wobj,bool cups{*},PERS loaddata load,num approachHeight)
        ! cups: cups on/off at the target, load: load after the target
        MoveJ Offs(target,0,0,approachHeight),TransitSpeed,z10,toolVacuum\WObj:=wobj;
        MoveL target,ApproachSpeed,fine,toolVacuum\WObj:=wobj;
        VacuumControl cups;
        GripLoad load;
        MoveL Offs(target,0,0,approachHeight),ApproachSpeed,z10,toolVacuum\WObj:=wobj;
    ENDPROC

    !-----------------------------------------------------------------------
    ! Calculation of approach heights (how much the robot goes up over the target)
    !-----------------------------------------------------------------------
    FUNC num ApproachHeight(num station)
        VAR num approachingHeight:=9E+09;
        TEST station
        CASE StationConveyor1:
            approachingHeight:=TransitHeight-ConveyorsHeight-Box1Height;
        CASE StationConveyor2:
            approachingHeight:=TransitHeight-ConveyorsHeight-Box2Height;
        CASE StationTable:
            approachingHeight:=TransitHeight-TableHeight-Box2Height;
        CASE StationLinerStand:
            approachingHeight:=TransitHeight-LinerStandHeight-linersLeft*LinerHeight;
        CASE StationHalfPallet:
            approachingHeight:=TransitHeight-HalfPalletHeight-HalfPalletLayerZ()-Box2Height-PalletOffsetHeight;
            IF approachingHeight<MinApproachHeight THEN
                approachingHeight:=MinApproachHeight;
            ENDIF
        CASE StationEuroPallet:
            approachingHeight:=TransitHeight-EuroPalletHeight-Box1Height*box1Layer-PalletOffsetHeight;
            IF approachingHeight<MinApproachHeight THEN
                approachingHeight:=MinApproachHeight;
            ENDIF
        DEFAULT:
            ! If another station is entered the robot will announce an error trying to reach 9E+09: Safety stop
        ENDTEST
        RETURN approachingHeight;
    ENDFUNC

    !-----------------------------------------------------------------------
    ! Assignment of logical cup signals with physical signals
    !-----------------------------------------------------------------------
    PROC InitSignals()
        ! Call it first: VacuumControl needs it
        AliasIO DO_Cup11,cupSignals{1};
        AliasIO DO_Cup12,cupSignals{2};
        AliasIO DO_Cup13,cupSignals{3};
        AliasIO DO_Cup21,cupSignals{4};
        AliasIO DO_Cup22,cupSignals{5};
        AliasIO DO_Cup23,cupSignals{6};
    ENDPROC

    !-----------------------------------------------------------------------
    ! Control of the vacuum of every cup
    !-----------------------------------------------------------------------
    PROC VacuumControl(bool cups{*})
        cupsState:=cups;

        FOR i FROM 1 TO Dim(cups,1) DO
            IF cups{i} THEN
                SetDO cupSignals{i},1;
            ELSE
                SetDO cupSignals{i},0;
            ENDIF
        ENDFOR

        ! Robot stopped in position, wait for the vacuum
        WaitTime\InPos,VacuumTime;
    ENDPROC

ENDMODULE

--- Controller Data/Controler/SYSPAR/EIO.cfg ---
EIO:CFG_1.0:6:1::
#
EIO_SIGNAL:

      -Name "DO_Cup11" -SignalType "DO" -Label "Vacuum valve gripper"\
      -Category "Gripper"

      -Name "DI_Box1Arrived" -SignalType "DI" -Label "Box 1 sensor conveyor 1"\
      -Category "Conveyor"

      -Name "DI_Box2Arrived" -SignalType "DI" -Label "Box 2 sensor conveyor 2"\
      -Category "Conveyor"

      -Name "DI_EuroPalletReplaced" -SignalType "DI"\
      -Label "Operator confirms new euro pallet" -Category "Operator"

      -Name "DI_HalfPalletReplaced" -SignalType "DI"\
      -Label "Operator confirms new half pallet" -Category "Operator"

      -Name "AI_VacuumPressure" -SignalType "AI"\
      -Label "Vacuum pressure sensor (bar)" -Category "Gripper" -MaxLog 10

      -Name "DO_Cup12" -SignalType "DO" -Label "Vacuum valve gripper"\
      -Category "Gripper"

      -Name "DO_Cup13" -SignalType "DO" -Label "Vacuum valve gripper"\
      -Category "Gripper"

      -Name "DO_Cup21" -SignalType "DO" -Label "Vacuum valve gripper"\
      -Category "Gripper"

      -Name "DO_Cup22" -SignalType "DO" -Label "Vacuum valve gripper"\
      -Category "Gripper"

      -Name "DO_Cup23" -SignalType "DO" -Label "Vacuum valve gripper"\
      -Category "Gripper"

      -Name "DI_LinersRefilled" -SignalType "DI"\
      -Label "Indicates refilled liners" -Category "Liners"

      -Name "DO_EuroPalletFull" -SignalType "DO"

      -Name "DO_HalfPalletFull" -SignalType "DO"

      -Name "DO_LinerStackEmpty" -SignalType "DO"
